(* IEC 61131-3 sources: POMIRTS_lab3/AS/Library/AsTCP, 3 files *)

(* ---- AsTCP.typ ---- *)
(********************************************************************
 * COPYRIGHT -- Bernecker + Rainer
 ********************************************************************
 * Library: AsTCP
 * File: AsTCP.typ
 * Author: B+R
 ********************************************************************
 * Data types of library AsTCP
 ********************************************************************)

TYPE
    tcpLINGER_typ		: STRUCT	(*linger*)
		lOnOff			: UDINT;	(*linger on/off*)
		lLinger			: UDINT;	(*linger time (seconds)*)
	END_STRUCT;

	tcpSO_ADDRESS_typ	: STRUCT	(*socket address*)
		pPort			: UDINT;	(*pointer where to store the portnumber*)
		pIpAddr			: UDINT;	(*pointer where to store the socket ip address*)
	END_STRUCT;
END_TYPE

(* ---- AsTCP.fun ---- *)
(********************************************************************
 * COPYRIGHT -- Bernecker + Rainer
 ********************************************************************
 * Library: AsTCP
 * File: AsTCP.fun
 * Author: B+R
 ********************************************************************
 * Functions and function blocks of library AsTCP
 ********************************************************************)

FUNCTION_BLOCK TcpOpen					(*opens a TCP socket; asynchronous execution*)
	VAR_INPUT
		enable			: BOOL;			(*enables execution*)
		pIfAddr			: UDINT;		(*pointer to the interface address*)
		port			: UINT;			(*port number of the socket*)
		options			: UDINT;		(*options that can be set during opening*)
	END_VAR

	VAR_OUTPUT
		status			: UINT;			(*execution status: ERR_OK, ERR_FUB_ENABLE_FALSE, ERR_FUB_BUSY, 0xXXXX = see help*)
		ident			: UDINT;		(*identifier for use with TcpServer, TcpClient, TcpSend, TcpRecv, TcpClose and TcpIoctl*)
	END_VAR

	VAR
        i_state			: UINT;			(*internal variable*)
		i_result		: UINT;			(*internal variable*)
        i_tmp			: UDINT;		(*internal variable*)
	END_VAR
END_FUNCTION_BLOCK

FUNCTION_BLOCK TcpServer				(*starts a TCP server; asynchronous execution*)
	VAR_INPUT
		enable			: BOOL;			(*enables execution*)
		ident			: UDINT;		(*identifier returned from TcpOpen()*)
		backlog			: UDINT;		(*number of connections to queue*)
		pIpAddr			: UDINT;		(*pointer where to store the ip address of the connected client*)
	END_VAR

	VAR_OUTPUT
		status			: UINT;			(*execution status: ERR_OK, ERR_FUB_ENABLE_FALSE, ERR_FUB_BUSY, 0xXXXX = see help*)
		identclnt		: UDINT;		(*identifier for use with fub TcpClose, TcpSend, and TcpRecv*)
		portclnt		: UINT;			(*port number of connected client*)
	END_VAR

	VAR
        i_state			: UINT;			(*internal variable*)
		i_result		: UINT;			(*internal variable*)
        i_tmp			: UDINT;		(*internal variable*)
	END_VAR
END_FUNCTION_BLOCK

FUNCTION_BLOCK TcpClient				(*establishs a connection to a TCP server; asynchronous execution*)
	VAR_INPUT
		enable			: BOOL;			(*enables execution*)
		ident			: UDINT;		(*identifier returned from TcpOpen()*)
		pServer			: UDINT;		(*pointer to the ip address of server to connect to*)
		portserv		: UINT;			(*port number of server to connect to*)
	END_VAR

	VAR_OUTPUT
		status			: UINT;			(*execution status: ERR_OK, ERR_FUB_ENABLE_FALSE, ERR_FUB_BUSY, 0xXXXX = see help*)
	END_VAR

	VAR
        i_state			: UINT;			(*internal variable*)
		i_result		: UINT;			(*internal variable*)
        i_tmp			: UDINT;		(*internal variable*)
	END_VAR
END_FUNCTION_BLOCK

FUNCTION_BLOCK TcpClose					(*closes a TCP socket and frees up all required resources; asynchronous execution*)
	VAR_INPUT
		enable			: BOOL;			(*enables execution*)
		ident			: UDINT;		(*identifier returned from TcpOpen()*)
		how				: UDINT;		(*shutdown behavior*)
	END_VAR

	VAR_OUTPUT
		status			: UINT;			(*execution status: ERR_OK, ERR_FUB_ENABLE_FALSE, ERR_FUB_BUSY, 0xXXXX = see help*)
	END_VAR

	VAR
        i_state			: UINT;			(*internal variable*)
		i_result		: UINT;			(*internal variable*)
        i_tmp			: UDINT;		(*internal variable*)
	END_VAR
END_FUNCTION_BLOCK

FUNCTION_BLOCK TcpSend					(*sends data (byte stream); asynchronous execution*)
	VAR_INPUT
		enable			: BOOL;			(*enables execution*)
		ident			: UDINT;		(*identifier returned from TcpOpen()*)
		pData			: UDINT;		(*pointer to the data to be sent*)
		datalen			: UDINT;		(*length of byte stream*)
		flags			: UDINT;		(*send flags (e.g. "out of band" data)*)
	END_VAR

	VAR_OUTPUT
		status			: UINT;			(*execution status: ERR_OK, ERR_FUB_ENABLE_FALSE, ERR_FUB_BUSY, 0xXXXX = see help*)
		sentlen			: UDINT;		(*number of actually sent bytes*)
	END_VAR

	VAR
        i_state			: UINT;			(*internal variable*)
		i_result		: UINT;			(*internal variable*)
        i_tmp			: UDINT;		(*internal variable*)
	END_VAR
END_FUNCTION_BLOCK

FUNCTION_BLOCK TcpRecv					(*receives TCP byte stream; asynchronous execution*)
	VAR_INPUT
		enable			: BOOL;			(*enables execution*)
		ident			: UDINT;		(*identifier returned from TcpOpen()*)
		pData			: UDINT;		(*pointer to the buffer where to store byte stream data*)
		datamax			: UDINT;		(*max. length of data in bytes*)
		flags			: UDINT;		(*receive flags*)
	END_VAR

	VAR_OUTPUT
		status			: UINT;			(*execution status: ERR_OK, ERR_FUB_ENABLE_FALSE, ERR_FUB_BUSY, 0xXXXX = see help*)
		recvlen			: UDINT;		(*length of the bytes received*)
	END_VAR

	VAR
        i_state			: UINT;			(*internal variable*)
		i_result		: UINT;			(*internal variable*)
        i_tmp			: UDINT;		(*internal variable*)
	END_VAR
END_FUNCTION_BLOCK

FUNCTION_BLOCK TcpIoctl					(*changes or retrieves settings; asynchronous execution*)
	VAR_INPUT
		enable			: BOOL;			(*enables execution*)
		ident			: UDINT;		(*identifier returned from TcpOpen()*)
		ioctl			: UDINT;		(*I/O control code*)
		pData			: UDINT;		(*pointer to the I/O control data buffer*)
		datalen			: UDINT;		(*lentgh of I/O control input data*)
	END_VAR

	VAR_OUTPUT
		status			: UINT;			(*execution status: ERR_OK, ERR_FUB_ENABLE_FALSE, ERR_FUB_BUSY, 0xXXXX = see help*)
		outlen			: UDINT;		(*output data length*)
	END_VAR

	VAR
        i_state			: UINT;			(*internal variable*)
		i_result		: UINT;			(*internal variable*)
        i_tmp			: UDINT;		(*internal variable*)
	END_VAR
END_FUNCTION_BLOCK

(* ---- AsTCP.var ---- *)
(********************************************************************
 * COPYRIGHT -- Bernecker + Rainer
 ********************************************************************
 * Library: AsTCP
 * File: AsTCP.var
 * Author: B+R
 ********************************************************************
 * Local variables of library AsTCP
 ********************************************************************)

VAR CONSTANT
	tcpERR_INVALID_IDENT				: UINT := 32600;	(*invalid ident*)
	tcpERR_NOMORE_IDENTS				: UINT := 32601;	(*no more idents*)
	tcpERR_ALREADY_EXIST				: UINT := 32602;	(*socket already exists*)
	tcpERR_PARAMETER					: UINT := 32603;	(*invalid parameter, check parameter*)
	tcpERR_INVALID_IOCTL				: UINT := 32604;	(*io control not supported*)
	tcpERR_NO_DATA						: UINT := 32605;	(*no data to receive*)
	tcpERR_SENTLEN						: UINT := 32606;	(*length sent error, call again*)
	tcpERR_WOULDBLOCK					: UINT := 32607;	(*would block, call again*)
	tcpERR_INVALID						: UINT := 32608;	(*invalid argument*)
	tcpERR_NOT_CONNECTED				: UINT := 32609;	(*socket is not connected*)
	tcpERR_ALREADY_CONNECTED			: UINT := 32610;	(*connected has been already established*)
	tcpERR_NO_OOBDATA					: UINT := 32611;	(*no out of band data*)
	tcpERR_INTERFACE					: UINT := 32612;	(*illegal interface*)
	tcpERR_NOCLIENT						: UINT := 32613;	(*client not yet connected*)

	tcpERR_SOCKET_CREATE				: UINT := 32650;	(*create socket failed*)
	tcpERR_SOCKET_BIND					: UINT := 32651;	(*bind socket failed*)
	tcpERR_SOCKET_LISTEN				: UINT := 32652;	(*listen socket failed*)
	tcpERR_SOCKET_ACCEPT				: UINT := 32653;	(*accept socket failed*)

	tcpERR_SYSTEM						: UINT := 32699;	(*system error*)

	tcpSO_LINGER_SET					: UDINT := 1001;	(*set option linger*)
	tcpSO_LINGER_GET					: UDINT := 1002;	(*get option linger*)
	tcpSO_KEEPALIVE_SET					: UDINT := 1003;	(*set option keep alive*)
	tcpSO_KEEPALIVE_GET					: UDINT := 1004;	(*get option keep alive*)
	tcpSO_SNDBUF_SET					: UDINT := 1005;	(*set option send buffer*)
	tcpSO_SNDBUF_GET					: UDINT := 1006;	(*get option send buffer*)
	tcpSO_RCVBUF_SET					: UDINT := 1007;	(*set option receive buffer*)
	tcpSO_RCVBUF_GET					: UDINT := 1008;	(*get option receive buffer*)
	tcpSO_OOBINLINE_SET					: UDINT := 1009;	(*set option out of band data inline*)
	tcpSO_OOBINLINE_GET					: UDINT := 1010;	(*get option out of band data inline*)
	tcpSO_ADDRESS_GET					: UDINT := 1011;	(*get socket address*)
	tcpSO_NOWAITING_SET					: UDINT := 1012;	(*set option no waiting until client connects*)
	tcpSO_NOWAITING_GET					: UDINT := 1013;	(*get option no waiting until client connects*)
	tcpTCP_NODELAY_SET					: UDINT := 2001;	(*set option tcp no delay*)
	tcpTCP_NODELAY_GET					: UDINT := 2002;	(*get option tcp no delay*)
	tcpID_LIST_GET						: UDINT := 3001;	(*get ident list*)
	tcpID_MAX_GET						: UDINT := 3002;	(*get max ident count*)

	tcpMSG_OOB							: UDINT := 1;		(*out of band message*)
	tcpMSG_PEEK							: UDINT := 2;		(*don't remove data from socket (receive)*)
	tcpMSG_DONTROUTE					: UDINT := 4;		(*message don't route (send)*)

	tcpOPT_REUSEADDR					: UDINT := 1;		(*option reuse address*)

	tcpSHUT_RD							: UDINT := 1;		(*shutdown read channel*)
	tcpSHUT_WR							: UDINT := 2;		(*shutdown write channel*)

	tcpINVALID_IDENT					: UDINT := 0;		(*invlaid ident*)
END_VAR
